(* PLC project g_independent_hp_trip_bomb, Anonymous Benchmark Suite 1.0 *)
(* stored: creationDateTime 2026-09-02T00:00:00 *)

PROGRAM g_independent_hp_trip_bomb
  VAR_INPUT
    pressure_high : BOOL;
    sequence_step_active : BOOL;
    maint : BOOL;
  END_VAR
  VAR_OUTPUT
    vent_valve : BOOL;
  END_VAR

(* LD diagram, written out as Structured Text *)
vent_valve := pressure_high AND (NOT maint OR sequence_step_active);
END_PROGRAM

CONFIGURATION Config0
  RESOURCE Res0 ON PLC
    TASK tcyclic(INTERVAL := T#10ms, PRIORITY := 0);
    PROGRAM inst0 WITH tcyclic : g_independent_hp_trip_bomb;
  END_RESOURCE
END_CONFIGURATION
